PROGRAM MAIN
VAR
	robot : RobotComposition;
END_VAR

robot.Execute();

END_PROGRAM

(* stored: Version 1.1.0.1, ProductVersion 3.1.4026.12
   POU MAIN: Id {6af6c587-617c-5902-b7b1-f003c23889d7}, SpecialFunc None *)
